Fanuc KAREL source: KT00233.KL

PROGRAM KT00233
%NOLOCKGROUP
VAR
  I1: INTEGER
  B2: BOOLEAN
  OUT: BOOLEAN
BEGIN
  I1 = 2
    B2 = FALSE
  OUT = I1 OR B2
END KT00233
